Yaskawa INFORM job: 12.JBI

/JOB
//NAME 12
//POS
///NPOS 25,25,25,0,0,0
///TOOL 0
///POSTYPE PULSE
///PULSE
C00000=-289,-101156,-84205,3690,-80188,-1943
C00001=-289,-101156,-84205,3690,-80188,-1943
C00002=85809,37752,10282,9567,-42392,-7198
C00003=91720,84357,22878,19424,-27586,-13450
C00004=92414,78654,15740,20967,-26356,-14358
C00005=92788,83783,22154,20355,-27669,-14125
C00006=92788,83472,22283,20198,-27894,-14045
C00007=93020,83548,21764,20611,-27608,-14298
C00008=92641,84026,22365,20234,-27644,-14035
C00009=92641,80164,24447,18310,-30735,-13050
C00010=93600,82568,20643,21184,-27565,-14699
C00011=93600,76074,24912,17799,-33205,-12945
C00012=94542,78896,16227,22502,-27005,-15543
C00013=94466,78056,15184,22601,-26793,-15578
C00014=94772,76457,13204,23142,-26501,-15912
C00015=95464,75690,12260,23823,-26497,-16391
C00016=95642,77087,13978,23685,-26850,-16360
C00017=94932,82677,20941,22097,-27988,-15422
C00018=96159,81404,19345,23236,-27978,-16238
C00019=96159,81404,19345,23236,-27978,-16238
C00020=96159,77644,21324,21134,-30905,-15159
C00021=97032,80203,17741,24144,-27852,-16869
C00022=97032,71197,24888,18870,-36288,-14091
C00023=-289,-101156,-84205,3690,-80188,-1943
C00024=-289,-101156,-84205,3690,-80188,-1943
BC00000=570125
BC00001=262324
BC00002=262818
BC00003=262818
BC00004=262818
BC00005=262818
BC00006=262818
BC00007=262818
BC00008=262818
BC00009=262818
BC00010=262818
BC00011=262818
BC00012=262818
BC00013=262818
BC00014=262818
BC00015=262818
BC00016=262818
BC00017=262818
BC00018=262818
BC00019=262818
BC00020=262818
BC00021=262818
BC00022=262818
BC00023=262324
BC00024=570125
EC00000=2713,0
EC00001=2713,0
EC00002=2712,0
EC00003=2712,0
EC00004=2712,0
EC00005=2712,0
EC00006=2712,0
EC00007=2712,0
EC00008=2712,0
EC00009=2712,0
EC00010=2712,0
EC00011=2712,0
EC00012=2712,0
EC00013=2712,0
EC00014=2712,0
EC00015=2712,0
EC00016=2712,0
EC00017=2712,0
EC00018=2712,0
EC00019=2712,0
EC00020=2712,0
EC00021=2712,0
EC00022=2712,0
EC00023=2713,0
EC00024=2713,0
//INST
///DATE 2019/11/16 12:30
///ATTR SC,RW
///GROUP1 RB1,BS1
///GROUP2 ST2
NOP
MOVJ C00000 BC00000 VJ=90.00  +MOVJ EC00000 VJ=90.00
MOVJ C00001 BC00001 VJ=90.00  +MOVJ EC00001 VJ=90.00
MOVJ C00002 BC00002 VJ=90.00  +MOVJ EC00002 VJ=90.00
MOVJ C00003 BC00003 VJ=90.00  +MOVJ EC00003 VJ=90.00
MACRO1 MJ#(0) ARGF1
ARCON
MOVL C00004 BC00004 V=5.0  +MOVJ EC00004 VJ=90.00
MOVL C00005 BC00005 V=5.0  +MOVJ EC00005 VJ=90.00
ARCOF
MOVJ C00006 BC00006 VJ=90.00  +MOVJ EC00006 VJ=90.00
MOVJ C00007 BC00007 VJ=90.00  +MOVJ EC00007 VJ=90.00
ARCON
MOVL C00008 BC00008 V=5.0  +MOVJ EC00008 VJ=90.00
ARCOF
MOVJ C00009 BC00009 VJ=90.00  +MOVJ EC00009 VJ=90.00
MOVJ C00010 BC00010 VJ=90.00  +MOVJ EC00010 VJ=90.00
ARCON
TIMER T=2.00
ARCOF
MOVJ C00011 BC00011 VJ=90.00  +MOVJ EC00011 VJ=90.00
MOVJ C00012 BC00012 VJ=90.00  +MOVJ EC00012 VJ=90.00
ARCON
MOVC C00013 BC00013 V=5.0  +MOVJ EC00013 VJ=90.00
MOVC C00014 BC00014 V=5.0  +MOVJ EC00014 VJ=90.00
MOVC C00015 BC00015 V=5.0  +MOVJ EC00015 VJ=90.00
MOVC C00016 BC00016 V=1350.0  +MOVJ EC00016 VJ=90.00
MOVL C00017 BC00017 V=5.0  +MOVJ EC00017 VJ=90.00
MOVJ C00018 BC00018 VJ=30.00  +MOVJ EC00018 VJ=90.00
MOVJ C00019 BC00019 VJ=30.00  +MOVJ EC00019 VJ=30.00
ARCOF
MOVJ C00020 BC00020 VJ=30.00  +MOVJ EC00020 VJ=30.00
MOVJ C00021 BC00021 VJ=30.00  +MOVJ EC00021 VJ=30.00
ARCON
TIMER T=2.00
ARCOF
MOVJ C00022 BC00022 VJ=30.00  +MOVJ EC00022 VJ=30.00
MOVJ C00023 BC00023 VJ=90.00  +MOVJ EC00023 VJ=90.00
MOVJ C00024 BC00024 VJ=90.00  +MOVJ EC00024 VJ=90.00
END
